# EPICS substitutions: db/Beckhoff_7XXX/ecmcEX72XX_OPT_cst.substitutions
file "ecmcEL72XX_DRV_CST.template"
{
  pattern {CH_ID, ESLO, EGU}
          {"$(OPT_CH_ID=01)", 0.1, "%"}
}
